FUNCTION_BLOCK AFIFO_UINT_TO_E (* Konverter: Socket AFIFO_UINT auf normale Events. DATA mit OUT/N kommt vom FIFO, PROCESSED geht ueber den Rueckkanal des Adapters an den FIFO zurueck. *)
  (* Standard: 61499-2; Description: Copyright (c) 2026 Meisterschulen am Ostbahnhof This program and the accompanying materials are made available under the terms of the Eclipse Public License 2.0 which is available at https://www.eclipse.org/legal/epl-2.0/ SPDX-License-Identifier: EPL-2.0 *)
  (* Version 1.0, 2026-11-08, Franz Höpfinger, Meisterschulen am Ostbahnhof, initial API and implementation and/or initial documentation *)
  PACKAGE FIFO_adapter;
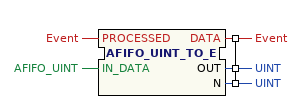
  EVENT_INPUT
    PROCESSED; (* Konsument bestaetigt: der zuletzt per DATA gelieferte Wert ist verarbeitet *)
  END_EVENT
  EVENT_OUTPUT
    DATA WITH OUT, N; (* Neuer Wert vom FIFO - es folgt kein weiteres DATA, bevor PROCESSED eingetroffen ist *)
  END_EVENT
  VAR_OUTPUT
    OUT : UINT; (* Gelieferter Wert *)
    N : UINT; (* Anzahl der danach noch wartenden Elemente in der Queue *)
  END_VAR
  SOCKETS
    IN_DATA : FIFO_adapter::AFIFO_UINT; (* Hier haengt der Plug OUT_DATA von FIFO_UINT_Adapter an *)
  END_SOCKETS
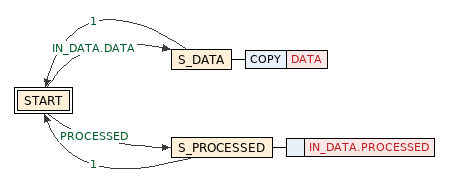
  EC_STATES
    START; (* Initial State *)
    S_DATA : COPY -> DATA;
    S_PROCESSED : -> IN_DATA.PROCESSED;
  END_STATES
  EC_TRANSITIONS
    START TO S_DATA := IN_DATA.DATA;
    S_DATA TO START := 1;
    START TO S_PROCESSED := PROCESSED;
    S_PROCESSED TO START := 1;
  END_TRANSITIONS
  ALGORITHM COPY IN ST: (* Wert und Fuellstand vom Adapter uebernehmen *)
OUT := IN_DATA.OUT;
N := IN_DATA.N;
  END_ALGORITHM
END_FUNCTION_BLOCK
